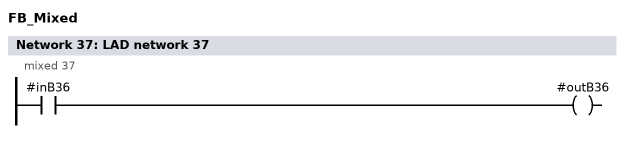
   RUNG wire#powerrail
      Contact( #inB36 )
      Coil( #outB36 )
   END_RUNG
   // the same network as SCL:
   #outB36 := #inB36;
END_REGION

REGION Network 38 (FBD): FBD network 38
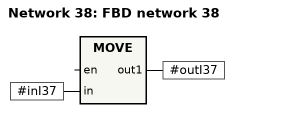
   #outI37 := #inI37;
END_REGION

REGION Network 39 (SCL): SCL network 39
   #tI38 := #inI38 + #cI8;
           IF #inB38 THEN
               #outR18 := #inR18 * 2.0;
           END_IF;
END_REGION

REGION Network 40: LAD network 40
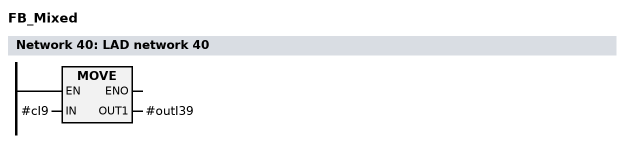
   RUNG wire#powerrail
      Move(in := #cI9, out1 => #outI39)
   END_RUNG
   // the same network as SCL:
   #outI39 := #cI9;
END_REGION

REGION Network 41 (FBD): FBD network 41
   // mixed 41
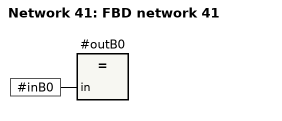
   #outB0 := #inB0;
END_REGION

REGION Network 42 (SCL): SCL network 42
   #tI41 := #inI1 + #cI11;
           IF #inB1 THEN
               #outR1 := #inR1 * 2.0;
           END_IF;
END_REGION

REGION Network 43: LAD network 43
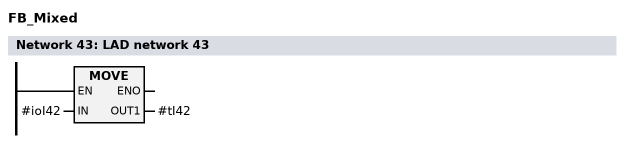
   RUNG wire#powerrail
      Move(in := #ioI42, out1 => #tI42)
   END_RUNG
   // the same network as SCL:
   #tI42 := #ioI42;
END_REGION

REGION Network 44 (FBD): FBD network 44
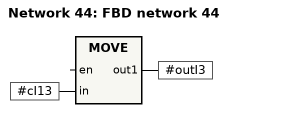
   #outI3 := #cI13;
END_REGION

REGION Network 45 (SCL): SCL network 45
   // mixed 45
   #tI44 := #inI4 + #cI14;
           IF #inB4 THEN
               #outR4 := #inR4 * 2.0;
           END_IF;
END_REGION

REGION Network 46: LAD network 46
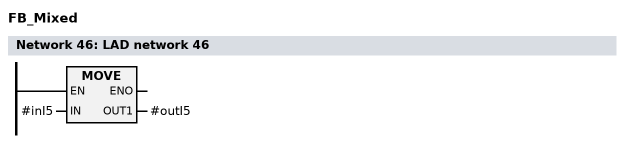
   RUNG wire#powerrail
      Move(in := #inI5, out1 => #outI5)
   END_RUNG
   // the same network as SCL:
   #outI5 := #inI5;
END_REGION

REGION Network 47 (FBD): FBD network 47
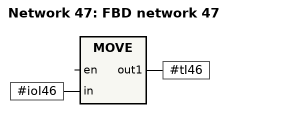
   #tI46 := #ioI46;
END_REGION

REGION Network 48 (SCL): SCL network 48
   #tI47 := #inI7 + #cI17;
           IF #inB7 THEN
               #outR7 := #inR7 * 2.0;
           END_IF;
END_REGION

REGION Network 49: LAD network 49
   // mixed 49
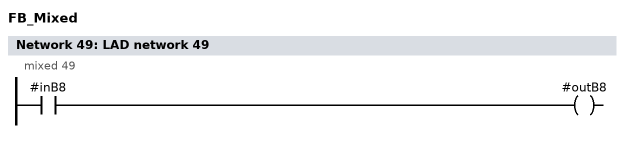
   RUNG wire#powerrail
      Contact( #inB8 )
      Coil( #outB8 )
   END_RUNG
   // the same network as SCL:
   #outB8 := #inB8;
END_REGION

REGION Network 50 (FBD): FBD network 50
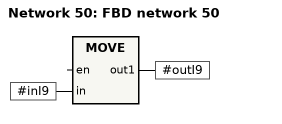
   #outI9 := #inI9;
END_REGION

REGION Network 51 (SCL): SCL network 51
   #tI50 := #inI10 + #cI20;
           IF #inB10 THEN
               #outR10 := #inR10 * 2.0;
           END_IF;
END_REGION

REGION Network 52: LAD network 52
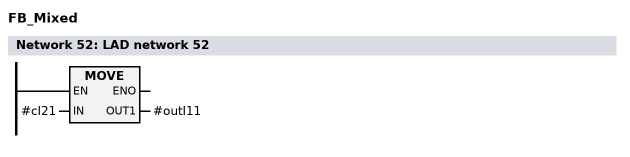
   RUNG wire#powerrail
      Move(in := #cI21, out1 => #outI11)
   END_RUNG
   // the same network as SCL:
   #outI11 := #cI21;
END_REGION

REGION Network 53 (FBD): FBD network 53
   // mixed 53
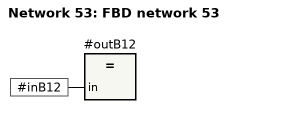
   #outB12 := #inB12;
END_REGION

REGION Network 54 (SCL): SCL network 54
   #tI53 := #inI13 + #cI23;
           IF #inB13 THEN
               #outR13 := #inR13 * 2.0;
           END_IF;
END_REGION

REGION Network 55: LAD network 55
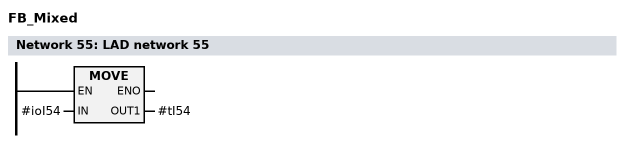
   RUNG wire#powerrail
      Move(in := #ioI54, out1 => #tI54)
   END_RUNG
   // the same network as SCL:
   #tI54 := #ioI54;
END_REGION

REGION Network 56 (FBD): FBD network 56
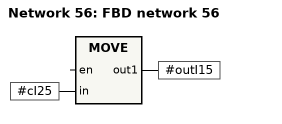
   #outI15 := #cI25;
END_REGION

REGION Network 57 (SCL): SCL network 57
   // mixed 57
   #tI56 := #inI16 + #cI26;
           IF #inB16 THEN
               #outR16 := #inR16 * 2.0;
           END_IF;
END_REGION

REGION Network 58: LAD network 58
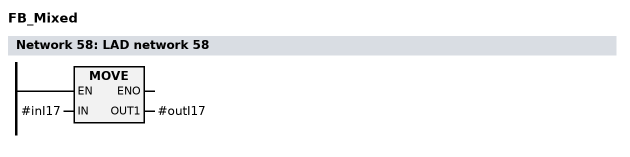
   RUNG wire#powerrail
      Move(in := #inI17, out1 => #outI17)
   END_RUNG
   // the same network as SCL:
   #outI17 := #inI17;
END_REGION

REGION Network 59 (FBD): FBD network 59
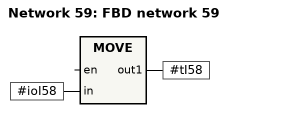
   #tI58 := #ioI58;
END_REGION

REGION Network 60 (SCL): SCL network 60
   #tI59 := #inI19 + #cI29;
           IF #inB19 THEN
               #outR19 := #inR19 * 2.0;
           END_IF;
END_REGION

REGION Network 61: LAD network 61
   // mixed 61
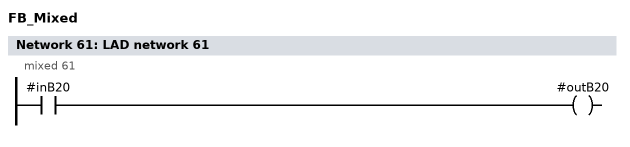
   RUNG wire#powerrail
      Contact( #inB20 )
      Coil( #outB20 )
   END_RUNG
   // the same network as SCL:
   #outB20 := #inB20;
END_REGION

REGION Network 62 (FBD): FBD network 62
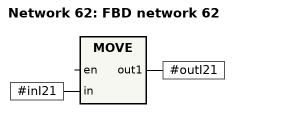
   #outI21 := #inI21;
END_REGION

REGION Network 63 (SCL): SCL network 63
   #tI62 := #inI22 + #cI2;
           IF #inB22 THEN
               #outR2 := #inR2 * 2.0;
           END_IF;
END_REGION

REGION Network 64: LAD network 64
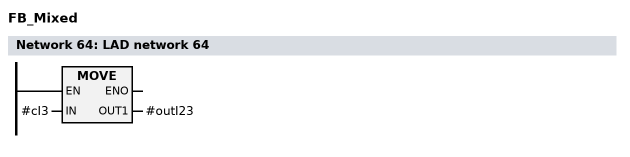
   RUNG wire#powerrail
      Move(in := #cI3, out1 => #outI23)
   END_RUNG
   // the same network as SCL:
   #outI23 := #cI3;
END_REGION

REGION Network 65 (FBD): FBD network 65
   // mixed 65
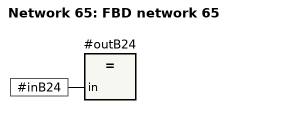
   #outB24 := #inB24;
END_REGION

REGION Network 66 (SCL): SCL network 66
   #tI65 := #inI25 + #cI5;
           IF #inB25 THEN
               #outR5 := #inR5 * 2.0;
           END_IF;
END_REGION

REGION Network 67: LAD network 67
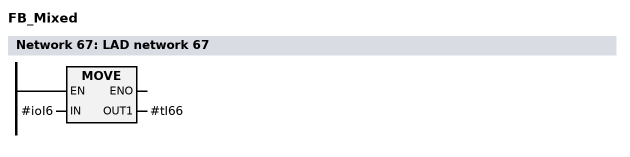
   RUNG wire#powerrail
      Move(in := #ioI6, out1 => #tI66)
   END_RUNG
   // the same network as SCL:
   #tI66 := #ioI6;
END_REGION

REGION Network 68 (FBD): FBD network 68
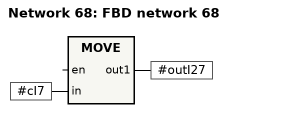
   #outI27 := #cI7;
END_REGION

REGION Network 69 (SCL): SCL network 69
   // mixed 69
   #tI68 := #inI28 + #cI8;
           IF #inB28 THEN
               #outR8 := #inR8 * 2.0;
           END_IF;
END_REGION

REGION Network 70: LAD network 70
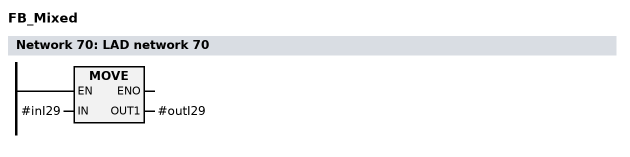
   RUNG wire#powerrail
      Move(in := #inI29, out1 => #outI29)
   END_RUNG
   // the same network as SCL:
   #outI29 := #inI29;
END_REGION

REGION Network 71 (FBD): FBD network 71
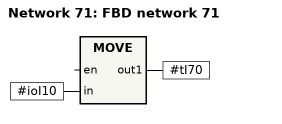
   #tI70 := #ioI10;
END_REGION

REGION Network 72 (SCL): SCL network 72
   #tI71 := #inI31 + #cI11;
           IF #inB31 THEN
               #outR11 := #inR11 * 2.0;
           END_IF;
END_REGION

REGION Network 73: LAD network 73
   // mixed 73
